(* IEC 61131-3 sources: JingjiangArm/moonboxpro_arm_8.4/Application/Application/任务列表/CommTask/RemoteEncSet, 4 files *)

(* ---- KS_CalcGCD.st ---- *)
(*@CES
Name=KS_CalcGCD
Type=FunctionBlock
TypeGuid=6f9dac99-8de1-4efc-8465-68ac443b7d08
Guid=2443a29b-db8f-4374-ad32-0269145bb8f6
HasDeclaration=True
HasImplementation=True
*)
{DECLARATION}
FUNCTION KS_CalcGCD : DWORD
(*计算最大公约数 by liu.yt*)
(*0代表未找到|出现死循环@最大10000*)
VAR_INPUT
	i_dwA:DWORD;
	i_dwB:DWORD;
END_VAR
VAR
	dwA:DWORD;
	dwB:DWORD;
	dwResult:DWORD;
	iCntNum:INT:=0;(*循环计数 防止死循环*)
	xNotFind: BOOL;
END_VAR

{IMPLEMENTATION}
dwA:=i_dwA;
dwB:=i_dwB;
IF (dwA = 0) THEN
	dwResult:=dwB;
ELSIF(dwB = 0) THEN
	dwResult:=dwB;
ELSE
	WHILE(dwB <> 0) DO
		dwResult:=dwB;
		dwB:=dwA MOD dwB;
		dwA:=dwResult;
		(*2025.12.11.172123+*)
		iCntNum:=iCntNum+1;
		IF iCntNum>=10000 THEN
			xNotFind:=TRUE;
			EXIT;
		END_IF
	END_WHILE
	(*未找到强制写0*)
	IF xNotFind THEN
		dwResult:=0;
	ELSE(*找到了*)
		dwResult:=dwA;
	END_IF
END_IF
KS_CalcGCD:=dwResult;

(* ---- KS_CheckDDA.st ---- *)
(*@CES
Name=KS_CheckDDA
Type=FunctionBlock
TypeGuid=6f9dac99-8de1-4efc-8465-68ac443b7d08
Guid=d0fb5f27-f5b4-42d1-b5c4-becbafc797f1
HasDeclaration=True
HasImplementation=True
*)
{DECLARATION}
FUNCTION KS_CheckDDA : BOOL(*false:DDA溢出@重新计算参数|TRUE:DDA正常*)
(*
检查dda处理的合法性@时钟运行周期时间内脉冲个数不能超过1.
获取到编码器值需要通过DDA插值处理,DDA插值的周期是时钟周期
如果时钟周期的脉冲变化量超过1,插值会出现丢失脉冲的情况
如果超过则输出不合法标志,并输出建议的编码器减速比(用于分频),编码器值@该值和库的计算公式有匹配关系
重新设置异站参数。
*)
(*
公式：dwDDAMotorEnc(DDA前分辨率)=i_dwMotorEncResolution*B/A
	  dwDDAMotorEnc(>> N@右移) = i_dwRemoteEnc
*)
(*i_dwRemoteEnc 该值是131072@和套色采样精度bit=>>5相关*)
VAR_INPUT
	i_byClock_MHZ			: BYTE:=125;(*时钟@mhz*)
	i_dwMotorEncResolution	: DWORD:=4194304;(*电机的编码器分辨率*)
	i_uiRotateSpeed_Max		: UINT:=3000;(*最大转速*)
	i_dwRemoteEnc			: DWORD:=131072;(*最终异站分辨率@131072|也是套色用的使用*)
	i_rMaxPulsePCycle		: REAL:=0.95;(*每个时钟周期最大脉冲数-不能超过1|目前125mhz即8ns的脉冲个数|适当小于1,留点余量*)
	i_puiA					: POINTER TO UINT;(*分母*)
	i_puiB					: POINTER TO UINT;(*分子*)
	i_pdwSetMotorEnc		: POINTER TO DWORD;(*设置的电机分辨率@目前等于输入的分辨率值*)
	i_pdwSetMotorEnc_DDA	: POINTER TO DWORD;(*DDA后电机分辨率@默认等于输入分辨率*)
	i_pbyRshBit				: POINTER TO BYTE;(*DDA后编码器右移位数*)
END_VAR
VAR
	iN					: INT;
	dwTmp				: DWORD;
	lrTmp				: LREAL;
	lrCoeff_Min2Ns		: LREAL;(*单位换算系数@MIN->ns*)
	byClock_ns			: BYTE;(*时间@ns*)
	rPulsePCycle		: REAL;(*每个周期的脉冲数*)
	rMaxPulsePCycle		: REAL;
	xOk					: BOOL;
	uiA					: UINT:=1;(*分母*)
	uiB					: UINT:=1;(*分子*)
	dwSetMotorEnc		: DWORD:=4194304;(*设置的电机分辨率*)
	byRshBit			: BYTE:=5;(*DDA后编码器右移位数@默认值*)
	dwDDAMotorEnc_Max	: DWORD;(*最大的dda编码器分辨率|*)
	dwDDAMotorEnc		: DWORD;(*可以用的@满足移位后的分辨率=131072*)
	dwSetMotorEnc_DDA	: DWORD;(*DDA后电机分辨率*)
	dwRemoteEnc			: DWORD:=131072;(*最终异站分辨率@131072*)
END_VAR

{IMPLEMENTATION}
(*获取单位周期脉冲的阈值*)
rMaxPulsePCycle:=i_rMaxPulsePCycle;
IF rMaxPulsePCycle>1 THEN
	rMaxPulsePCycle:=1;
END_IF
(*获取异站的最终分辨率*)
dwRemoteEnc:=i_dwRemoteEnc;
IF dwRemoteEnc=0 THEN
	dwRemoteEnc:=131072;
END_IF
(*周期时间计算*)
IF i_byClock_MHZ<>0 THEN
	lrTmp:=1000.0 / BYTE_TO_LREAL(i_byClock_MHZ) ;(*ns*)
ELSE
	lrTmp:=8;
END_IF
byClock_ns:=LREAL_TO_BYTE(lrTmp);(*周期@ns*)
(*单位周期的脉冲数*)
lrCoeff_Min2Ns:=60.0 * 1000 * 1000 * 1000;
lrTmp:=UINT_TO_LREAL(i_uiRotateSpeed_Max) * i_dwMotorEncResolution;(*脉冲p/min*)
lrTmp:=lrTmp / lrCoeff_Min2Ns;(*脉冲/ns*)
lrTmp:=lrTmp * byClock_ns;(*单位周期的脉冲数*)
rPulsePCycle:=lrTmp;
(*阈值判断*)
IF rPulsePCycle <= rMaxPulsePCycle THEN(*正常*)
	xOk:=TRUE;
ELSE(*脉冲太快了*)
	xOk:=FALSE;
	rPulsePCycle:=rMaxPulsePCycle;(*每个周期的脉冲按照最大值|用于反算参数@pulse/ns*)
END_IF
(*计算建议的分频值和配置的分辨率值*)
dwSetMotorEnc:=i_dwMotorEncResolution;
dwSetMotorEnc_DDA:=dwSetMotorEnc;
IF NOT xOk THEN
	(*重新计算设置值*)
	(*反算DDA前输入的电机分辨率*)
	lrTmp:=rPulsePCycle / byClock_ns;(*单位p/ns*)
	lrTmp:=lrTmp * lrCoeff_Min2Ns;(*单位p/min*)
	lrTmp:=lrTmp / i_uiRotateSpeed_Max;(*单位p/r@即可以用的最大电机的分辨率*)
	dwDDAMotorEnc_Max:=LREAL_TO_DWORD(lrTmp);(*写入到dword*)

	(*DDA输入的分辨率经过变比(>>N@右移)需要=dwRemoteEnc|反算改变比*)
	dwTmp:= dwDDAMotorEnc_Max / dwRemoteEnc;(*保留整数*)
	(*未找到以2为低的对数公式|用循环找吧*)
	FOR iN:=2 TO 20 BY 1 DO(*最大右移20*)
		lrTmp:=EXPT(2,iN);(*2的n次方*)
		IF lrTmp > dwTmp THEN(*超过了倍数|取上一个*)
			iN:=iN-1;
			EXIT;
		ELSIF lrTmp = dwTmp THEN(*找到了*)
			EXIT;
		END_IF
	END_FOR
	byRshBit:=INT_TO_BYTE(iN);(*2025.12.9.193202*)
	dwDDAMotorEnc:=REAL_TO_DWORD(dwRemoteEnc * EXPT(2,iN));(*反算出进入dda的电机分辨率*)
	(*使用实际分辨率计算ab*)
	dwTmp:=KS_CalcGCD(dwDDAMotorEnc,i_dwMotorEncResolution);(*计算最大共约数*)
	IF dwTmp<>0 THEN
		uiA := DWORD_TO_UINT(i_dwMotorEncResolution / dwTmp);
		uiB := DWORD_TO_UINT(dwDDAMotorEnc / dwTmp);
	ELSE
		uiA:=1;
		uiB:=1;
	END_IF
	dwSetMotorEnc_DDA:=dwDDAMotorEnc;(*输出dda后的电机分辨率*)
END_IF
IF i_puiA<>0 THEN
	i_puiA^:=uiA;
END_IF
IF i_puiB<>0 THEN
	i_puiB^:=uiB;
END_IF
IF i_pdwSetMotorEnc<>0 THEN
	i_pdwSetMotorEnc^:=dwSetMotorEnc;
END_IF
IF i_pdwSetMotorEnc_DDA<>0 THEN
	i_pdwSetMotorEnc_DDA^:=dwSetMotorEnc_DDA;
END_IF
IF i_pbyRshBit<>0 THEN
	i_pbyRshBit^:=byRshBit;
END_IF
KS_CheckDDA:=xOk;

(* ---- KS_GetRemoteEncParam.st ---- *)
(*@CES
Name=KS_GetRemoteEncParam
Type=FunctionBlock
TypeGuid=6f9dac99-8de1-4efc-8465-68ac443b7d08
Guid=5c03e2a5-041e-48c9-9983-827936801836
HasDeclaration=True
HasImplementation=True
*)
{DECLARATION}
FUNCTION KS_GetRemoteEncParam : BOOL
VAR_INPUT
	i_xGet:BOOL;
	i_byStationId:BYTE;
	i_puiA:POINTER TO UINT;
	i_puiB:POINTER TO UINT;
	i_puiN:POINTER TO UINT;
	i_dwMotorEnc:POINTER TO DWORD;
	i_dwMotorEnc_DDA:POINTER TO DWORD;
END_VAR
VAR
	diTmp:DINT;
END_VAR

{IMPLEMENTATION}
IF i_xGet THEN
	(*DDA后移位N*)
	GT_RN_UserRemoteEncRd(0,ADR(diTmp),i_byStationId);
	IF i_puiN<>0 THEN
		i_puiN^:=DINT_TO_UINT(diTmp);
	END_IF
	(*DDA后编码器分辨率*)
	GT_RN_UserRemoteEncRd(1,ADR(diTmp),i_byStationId);
	IF i_puiN<>0 THEN
		i_dwMotorEnc_DDA^:=DINT_TO_DWORD(diTmp);
	END_IF
	(*电机编码器分辨率*)
	GT_RN_UserRemoteEncRd(2,ADR(diTmp),i_byStationId);
	IF i_puiN<>0 THEN
		i_dwMotorEnc^:=DINT_TO_DWORD(diTmp);
	END_IF

	(*设置减速比A*)
	GT_RN_UserRemoteEncRd(3,ADR(diTmp),i_byStationId);
	IF i_puiA<>0 THEN
		i_puiA^:=DINT_TO_UINT(diTmp);
	END_IF

	(*设置减速比b*)
	GT_RN_UserRemoteEncRd(4,ADR(diTmp),i_byStationId);
	IF i_puiB<>0 THEN
		i_puiB^:=DINT_TO_UINT(diTmp);
	END_IF

END_IF

(* ---- KS_SetRemoteEncParam.st ---- *)
(*@CES
Name=KS_SetRemoteEncParam
Type=FunctionBlock
TypeGuid=6f9dac99-8de1-4efc-8465-68ac443b7d08
Guid=52359865-76ae-4a72-8575-b7942d579f0c
HasDeclaration=True
HasImplementation=True
*)
{DECLARATION}
FUNCTION KS_SetRemoteEncParam : INT(*异站设置函数@用于月光系列*)
(*月光宝盒异站编码器设置功能@pro也使用*)
(*<0 代表设置失败*)
(*再次设置需要复位设置完成和设置失败标志*)
(*目前异站公式解释@仅代表2025.12.4时*)
(*
异站编码器输出必须是131072,
公式是 (输入编码器分辨率 * b / a)-> DDA ->DDA后分辨率 >> n = 131072
分辨率太大,或者减速比设置不合适会引起DDA处理溢出
DDA:按照125M(8ns)进行插值,不溢出原则是8ns时间编码器值不能>1
*)
VAR_INPUT
	i_xUseLocalEnc:BOOL;(*使用本地编码器*)
	i_iStationId:INT;(*站号@月光宝盒的*)
	i_dwMotorEncResolution:DWORD;(*电机的编码器分辨率*)
	i_uiRotateSpeed_Max:UINT;(*最大转速*)
	i_dwRemoteEnc: DWORD:=131072;(*最终异站分辨率@131072|也是套色用的使用*)
	i_pxSetDne:POINTER TO BOOL;(*设置完成*)
	i_pxSetFailed:POINTER TO BOOL;(*设置失败*)
END_VAR
VAR
	xSetDne:BOOL;(*设置完成*)
	xSetFailed:BOOL;(*设置完成*)
	iRtn: INT;
	xUpdateRtn: BOOL;(*更新返回值*)
	byStationId:BYTE;
	uiA: UINT;
	uiB: UINT;
	dwSetMotorEnc: DWORD;
	dwRemoteEnc: DWORD:=131072;(*最终异站分辨率@131072|也是套色用的使用*)
	dwSetMotorEnc_DDA	: DWORD;(*DDA后电机分辨率*)
	byRshBit			: BYTE:=5;(*DDA后编码器右移位数*)
	byUseLocalEnc		: BYTE;
	sTemp : STRING;
	uitime:UINT:=15225;(*临时测试，不需要同步*)

END_VAR
{IMPLEMENTATION}
IF i_pxSetDne<>0 THEN
	xSetDne:=i_pxSetDne^;
END_IF
IF i_pxSetFailed<>0 THEN
	xSetFailed:=i_pxSetFailed^;
END_IF
dwRemoteEnc:=i_dwRemoteEnc;(*2025.12.9.192118+*)
IF dwRemoteEnc=0 THEN
	dwRemoteEnc:=131072;
END_IF
sTemp := '';
IF (NOT xSetDne) OR (NOT xSetFailed) THEN

	IF i_iStationId>=0 AND i_iStationId<USER_MAX_STATION_NUM_V1 THEN
		byStationId:=INT_TO_BYTE(i_iStationId);
		(*检查dda是否过速度*)
		KS_CheckDDA(
			125(*i_byClock_MHZ*),
			i_dwMotorEncResolution(*i_dwMotorEncResolution*),
			i_uiRotateSpeed_Max(*i_uiRotateSpeed_Max*),
			dwRemoteEnc(*i_dwRemoteEnc*),
			0.95(*i_rMaxPulsePCycle*),
			ADR(uiA)(*i_puiA*),
			ADR(uiB)(*i_puiB*),
			ADR(dwSetMotorEnc)(*i_pdwSetMotorEnc*),
			ADR(dwSetMotorEnc_DDA)(*i_pdwSetMotorEnc_DDA*),
			ADR(byRshBit)(*i_pbyRshBit*));
		(*异站参数配置*)
		(*设置dda后右移位数*)
		//iRtn:=GT_RN_UserRemoteEncWr(0,byRshBit,byStationId);
		iRtn := GTN_RN_SetCameraRemoteEncParam(
			cardIndex:= 1,
			busIndex:= 1,
			stationPhyId:= byStationId,
			encIndex:= 0,
			paramIndex:= 0,
			paramValue:= byRshBit);

			sTemp := CONCAT(' StationId: ',BYTE_TO_STRING(byStationId));
			sTemp := CONCAT(sTemp,' byRshBit: ');
			sTemp := CONCAT(sTemp,BYTE_TO_STRING(byRshBit));
			sTemp := CONCAT(sTemp,' iRtn: ');
			KS_HY_AddMsgToLog(g_pstStHYLogFifo, LOG_LEVEL_DEBUG,sTemp, INT_TO_STRING(iRtn));
		IF iRtn=0 THEN(*设置正常*)
			(*设置经过变比后的dda分辨率*)
			//iRtn:=GT_RN_UserRemoteEncWr(1,dwSetMotorEnc_DDA,byStationId);
			iRtn := GTN_RN_SetCameraRemoteEncParam(
				cardIndex:= 1,
				busIndex:= 1,
				stationPhyId:= byStationId,
				encIndex:= 0,
				paramIndex:= 1,
				paramValue:= dwSetMotorEnc_DDA);

			sTemp := CONCAT(' StationId: ',BYTE_TO_STRING(byStationId));
			sTemp := CONCAT(sTemp,' dwSetMotorEnc_DDA: ');
			sTemp := CONCAT(sTemp,DWORD_TO_STRING(dwSetMotorEnc_DDA));
			sTemp := CONCAT(sTemp,' iRtn: ');
			KS_HY_AddMsgToLog(g_pstStHYLogFifo, LOG_LEVEL_DEBUG,sTemp, INT_TO_STRING(iRtn));
		END_IF
		IF iRtn=0 THEN(*设置正常*)
			(*设置电机实际分辨率*)
			//iRtn:=GT_RN_UserRemoteEncWr(2,dwSetMotorEnc,byStationId);
			iRtn := GTN_RN_SetCameraRemoteEncParam(
				cardIndex:= 1,
				busIndex:= 1,
				stationPhyId:= byStationId,
				encIndex:= 0,
				paramIndex:= 2,
				paramValue:= dwSetMotorEnc);
	//2026.5.12.164334
			sTemp := CONCAT(' StationId: ',BYTE_TO_STRING(byStationId));
			sTemp := CONCAT(sTemp,' dwSetMotorEnc: ');
			sTemp := CONCAT(sTemp,DWORD_TO_STRING(dwSetMotorEnc));
			sTemp := CONCAT(sTemp,' iRtn: ');
			KS_HY_AddMsgToLog(g_pstStHYLogFifo, LOG_LEVEL_DEBUG,sTemp, INT_TO_STRING(iRtn));
		END_IF
		IF iRtn=0 THEN(*设置正常*)
			(*设置变比a*)
			//iRtn:=GT_RN_UserRemoteEncWr(3,uiA,byStationId);
			iRtn := GTN_RN_SetCameraRemoteEncParam(
				cardIndex:= 1,
				busIndex:= 1,
				stationPhyId:= byStationId,
				encIndex:= 0,
				paramIndex:= 3,
				paramValue:= uiA);
//2026.5.12.164330
			sTemp := CONCAT(' StationId: ',BYTE_TO_STRING(byStationId));
			sTemp := CONCAT(sTemp,' uiA: ');
			sTemp := CONCAT(sTemp,UINT_TO_STRING(uiA));
			sTemp := CONCAT(sTemp,' iRtn: ');
			KS_HY_AddMsgToLog(g_pstStHYLogFifo, LOG_LEVEL_DEBUG,sTemp, INT_TO_STRING(iRtn));
		END_IF
		IF iRtn=0 THEN(*设置正常*)
			(*设置变比b*)
			//iRtn:=GT_RN_UserRemoteEncWr(4,uiB,byStationId);
			iRtn := GTN_RN_SetCameraRemoteEncParam(
				cardIndex:= 1,
				busIndex:= 1,
				stationPhyId:= byStationId,
				encIndex:= 0,
				paramIndex:= 4,
				paramValue:= uiB);

			sTemp := CONCAT(' StationId: ',BYTE_TO_STRING(byStationId));
			sTemp := CONCAT(sTemp,' uiB: ');
			sTemp := CONCAT(sTemp,UINT_TO_STRING(uiB));
			sTemp := CONCAT(sTemp,' iRtn: ');
			KS_HY_AddMsgToLog(g_pstStHYLogFifo, LOG_LEVEL_DEBUG,sTemp, INT_TO_STRING(iRtn));
		END_IF
		(*2026.05.13.103437临时测试，不需要同步*)
		IF iRtn=0 THEN(*设置正常*)
			(*设置变比a*)
			//iRtn:=GT_RN_UserRemoteEncWr(3,uiA,byStationId);
			iRtn := GTN_RN_SetCameraRemoteEncParam(
				cardIndex:= 1,
				busIndex:= 1,
				stationPhyId:= byStationId,
				encIndex:= 0,
				paramIndex:= 7,
				paramValue:= uitime);

		END_IF

		IF iRtn=0 THEN(*设置正常*)
			(*设置为异站或者本地*)
			IF i_xUseLocalEnc THEN(*本地*)
				byUseLocalEnc:=0;
			ELSE
				byUseLocalEnc:=1;
			END_IF
			//iRtn:=GT_RN_SetYGBHRemoteEnable(byUseLocalEnc,byStationId);(*TRUE:异站|FALSE:本地*)
			iRtn := GTN_RN_SetYGBHRemoteEnable(cardIndex:= 1, busIndex:= 1, enable:= byUseLocalEnc, station_id:= byStationId);

			sTemp := CONCAT(' StationId: ',BYTE_TO_STRING(byStationId));
			sTemp := CONCAT(sTemp,' byUseLocalEnc: ');
			sTemp := CONCAT(sTemp,BYTE_TO_STRING(byUseLocalEnc));
			sTemp := CONCAT(sTemp,' iRtn: ');
			KS_HY_AddMsgToLog(g_pstStHYLogFifo, LOG_LEVEL_DEBUG,sTemp, INT_TO_STRING(iRtn));
		END_IF

		IF iRtn=0 THEN(*设置正常*)
			xSetDne:=TRUE;
		ELSE
			xSetFailed:=TRUE;
		END_IF
		xUpdateRtn:=TRUE;
	END_IF
ELSE;
END_IF
IF i_pxSetDne<>0 THEN
	i_pxSetDne^:=xSetDne;
END_IF
IF i_pxSetFailed<>0 THEN
	i_pxSetFailed^:=xSetFailed;
END_IF

IF xUpdateRtn THEN
	KS_SetRemoteEncParam:=iRtn;
END_IF
